(* IEC 61131-3 sources: plc-st-coding-agent/progress/evidence/f14_v10_full_20261113/jobs/codex_minimax-m27 (part 8) *)

(* ---- self-medium-03.raw_candidate_04.st ---- *)
TYPE EState :
    (
        IDLE    := 0,
        OPENING := 1,
        CLOSING := 2,
        FAULT   := 3
    )
END_TYPE

FUNCTION_BLOCK FB
VAR_INPUT
    openBtn    : BOOL;
    closeBtn   : BOOL;
    openLimit  : BOOL;
    closeLimit : BOOL;
    obstacle   : BOOL;
END_VAR
VAR_OUTPUT
    motorUp    : BOOL;
    motorDown  : BOOL;
    errorFlag  : BOOL;
END_VAR
VAR
    state          : EState := IDLE;
    prev_openBtn   : BOOL := FALSE;
    prev_closeBtn  : BOOL := FALSE;
    prev_obstacle  : BOOL := FALSE;
    openRTrig      : R_TRIG;
    closeRTrig     : R_TRIG;
    dualRTrig      : R_TRIG;
END_VAR

(*
ENGINEERING_CONTRACT
===================
| Output/State | Activation           | Retention           | Reset/Deactivation              | Scan Priority | Units   |
|--------------|----------------------|---------------------|----------------------------------|---------------|---------|
| motorUp      | IDLE+rising(openBtn) | Running continues   | obstacle/openLimit/FAULT         | Same-scan     | BOOL    |
| motorDown    | IDLE+rising(closeBtn)| Running continues   | obstacle/closeLimit/FAULT        | Same-scan     | BOOL    |
| errorFlag    | Any state+obstacle   | Latched in FAULT    | No obstacle+dualBtn rising edge  | Highest       | BOOL    |
| state=FAULT  | Any state+obstacle   | Until dualBtn reset | No obstacle+dualBtn rising edge  | Highest       | EState  |
| state=IDLE   | Power-on/limit/reset | Until rising edge   | -                                | Default       | EState  |
PUB001: power-on IDLE
PUB002: init FALSE
PUB003-005: no obstacle IDLE start (openBtn rising, closeBtn=FALSE, not openLimit)
PUB006: dual-btn does not start
PUB007: motor command same-scan on start
PUB008-009: button release / direction buttons ignored during movement
PUB010-011: limit stop same-scan, opposite limit irrelevant
PUB012: mutual exclusion always
PUB013-014: obstacle → both stop + FAULT (highest priority)
PUB017-018: errorFlag latched, motors stopped in FAULT
PUB019-021: reset requires no obstacle + dualBtn from not-both to both
PUB022-024: reset → IDLE, same-scan stop, then follow rule 1
*)

BEGIN
    openRTrig(CLK := openBtn);
    closeRTrig(CLK := closeBtn);
    dualRTrig(CLK := openBtn AND closeBtn);

    (* Priority 1: Obstacle → immediate both-stop + FAULT *)
    IF obstacle THEN
        motorUp   := FALSE;
        motorDown := FALSE;
        state     := FAULT;
        errorFlag := TRUE;
    ELSE
        CASE state OF
            IDLE:
                motorUp   := FALSE;
                motorDown := FALSE;
                (* Start opening: rising edge of openBtn, closeBtn=FALSE, not at openLimit *)
                IF openRTrig.Q AND NOT closeBtn AND NOT openLimit THEN
                    motorUp := TRUE;
                    state   := OPENING;
                (* Start closing: rising edge of closeBtn, openBtn=FALSE, not at closeLimit *)
                ELSIF closeRTrig.Q AND NOT openBtn AND NOT closeLimit THEN
                    motorDown := TRUE;
                    state     := CLOSING;
                END_IF;

            OPENING:
                motorUp   := TRUE;
                motorDown := FALSE;
                IF openLimit THEN
                    motorUp := FALSE;
                    state   := IDLE;
                END_IF;

            CLOSING:
                motorUp   := FALSE;
                motorDown := TRUE;
                IF closeLimit THEN
                    motorDown := FALSE;
                    state     := IDLE;
                END_IF;

            FAULT:
                motorUp   := FALSE;
                motorDown := FALSE;
                IF dualRTrig.Q THEN
                    errorFlag := FALSE;
                    state     := IDLE;
                END_IF;
        END_CASE;
    END_IF;

    prev_openBtn  := openBtn;
    prev_closeBtn := closeBtn;
    prev_obstacle := obstacle;
END_FUNCTION_BLOCK

(* CONTRACT_RULES [] *)

(* ---- self-medium-04.candidate_01.st ---- *)
(* ENGINEERING_CONTRACT
 * Filling Valve Controller - Discrete Scan State Machine
 *
 * | State            | Activation           | Retention           | Explicit Reset       | Same-scan Priority | Units/Boundaries     |
 * |------------------|----------------------|---------------------|----------------------|--------------------|----------------------|
 * | valveOpen=FALSE  | resetBtn rising      | N/A (output only)   | N/A                  | highest            | BOOL                 |
 * | valveOpen=TRUE   | rising(startBtn) & !prev(valveOpen) | while accVol < targetVol | resetBtn rising | 2nd            | accumulated REAL [0, ∞) |
 * | pendingFill=TRUE | valve closes (accVol>=target) | until doneSensor=TRUE OR new start OR reset | resetBtn rising | 3rd            | BOOL internal state       |
 * | fillsToday++     | doneSensor=TRUE & pendingFill | N/A (output only)  | resetBtn rising      | lowest             | INT [0..32767]           |
 *
 * PUB002: startBtn rising edge detection uses prevStartBtn
 * PUB003: resetBtn rising edge detection uses prevResetBtn
 * PUB004: doneSensor read as level each scan (PUB004)
 * PUB005: flowVol added each scan including start scan
 * PUB006: accumulated >= targetVol triggers valve close same scan
 * PUB007: doneSensor checked immediately after valve close
 * PUB008: if doneSensor=TRUE same scan, confirm and clear pendingFill
 * PUB009: if doneSensor=FALSE, pendingFill retained for later confirmation
 * PUB010: fillsToday increments by 1 per confirmation
 * PUB011: fillsToday saturates at 32767
 * PUB012: resetBtn rising clears all state (valveOpen, accumulatedVol, pendingFill, fillsToday)
 * PUB035: new start cancels pendingFill immediately
 * PUB043: continuous doneSensor=TRUE does not double-count
 *)
FUNCTION_BLOCK FB
VAR_INPUT
    startBtn    : BOOL;
    resetBtn    : BOOL;
    doneSensor  : BOOL;
    targetVol   : REAL;
    flowVol     : REAL;
END_VAR
VAR_OUTPUT
    valveOpen   : BOOL := FALSE;
    fillsToday  : INT  := 0;
END_VAR
VAR
    prevStartBtn    : BOOL := FALSE;
    prevResetBtn    : BOOL := FALSE;
    accumulatedVol  : REAL := 0.0;
    pendingFill     : BOOL := FALSE;
END_VAR

    // Priority 1: Reset clears everything, no other action this scan
    IF resetBtn AND NOT prevResetBtn THEN
        valveOpen       := FALSE;
        accumulatedVol  := 0.0;
        pendingFill     := FALSE;
        fillsToday      := 0;
        prevStartBtn    := startBtn;
        prevResetBtn    := resetBtn;
        RETURN;
    END_IF;

    // Priority 2: Start new bottle (clears any pending confirmation)
    IF startBtn AND NOT prevStartBtn THEN
        pendingFill    := FALSE;
        accumulatedVol := 0.0;
        valveOpen      := TRUE;
        // flowVol added in filling section below
    END_IF;

    // Priority 3: Filling state - accumulate flow and check target
    IF valveOpen THEN
        accumulatedVol := accumulatedVol + flowVol;
        IF accumulatedVol >= targetVol THEN
            valveOpen := FALSE;
            // Immediate doneSensor check after valve close
            IF doneSensor THEN
                pendingFill := FALSE;
                IF fillsToday < 32767 THEN
                    fillsToday := fillsToday + 1;
                END_IF;
            ELSE
                pendingFill := TRUE;
            END_IF;
        END_IF;
    END_IF;

    // Priority 4: Pending confirmation - wait for doneSensor
    IF pendingFill AND doneSensor THEN
        pendingFill := FALSE;
        IF fillsToday < 32767 THEN
            fillsToday := fillsToday + 1;
        END_IF;
    END_IF;

    prevStartBtn := startBtn;
    prevResetBtn := resetBtn;
END_FUNCTION_BLOCK

(* CONTRACT_RULES [] *)

(* ---- self-medium-04.raw_candidate_01.st ---- *)
(* ENGINEERING_CONTRACT
 * Filling Valve Controller - Discrete Scan State Machine
 *
 * | State            | Activation           | Retention           | Explicit Reset       | Same-scan Priority | Units/Boundaries     |
 * |------------------|----------------------|---------------------|----------------------|--------------------|----------------------|
 * | valveOpen=FALSE  | resetBtn rising      | N/A (output only)   | N/A                  | highest            | BOOL                 |
 * | valveOpen=TRUE   | rising(startBtn) & !prev(valveOpen) | while accVol < targetVol | resetBtn rising | 2nd            | accumulated REAL [0, ∞) |
 * | pendingFill=TRUE | valve closes (accVol>=target) | until doneSensor=TRUE OR new start OR reset | resetBtn rising | 3rd            | BOOL internal state       |
 * | fillsToday++     | doneSensor=TRUE & pendingFill | N/A (output only)  | resetBtn rising      | lowest             | INT [0..32767]           |
 *
 * PUB002: startBtn rising edge detection uses prevStartBtn
 * PUB003: resetBtn rising edge detection uses prevResetBtn
 * PUB004: doneSensor read as level each scan (PUB004)
 * PUB005: flowVol added each scan including start scan
 * PUB006: accumulated >= targetVol triggers valve close same scan
 * PUB007: doneSensor checked immediately after valve close
 * PUB008: if doneSensor=TRUE same scan, confirm and clear pendingFill
 * PUB009: if doneSensor=FALSE, pendingFill retained for later confirmation
 * PUB010: fillsToday increments by 1 per confirmation
 * PUB011: fillsToday saturates at 32767
 * PUB012: resetBtn rising clears all state (valveOpen, accumulatedVol, pendingFill, fillsToday)
 * PUB035: new start cancels pendingFill immediately
 * PUB043: continuous doneSensor=TRUE does not double-count
 *)
FUNCTION_BLOCK FB
VAR_INPUT
    startBtn    : BOOL;
    resetBtn    : BOOL;
    doneSensor  : BOOL;
    targetVol   : REAL;
    flowVol     : REAL;
END_VAR
VAR_OUTPUT
    valveOpen   : BOOL := FALSE;
    fillsToday  : INT  := 0;
END_VAR
VAR
    prevStartBtn    : BOOL := FALSE;
    prevResetBtn    : BOOL := FALSE;
    accumulatedVol  : REAL := 0.0;
    pendingFill     : BOOL := FALSE;
END_VAR

    // Priority 1: Reset clears everything, no other action this scan
    IF resetBtn AND NOT prevResetBtn THEN
        valveOpen       := FALSE;
        accumulatedVol  := 0.0;
        pendingFill     := FALSE;
        fillsToday      := 0;
        prevStartBtn    := startBtn;
        prevResetBtn    := resetBtn;
        RETURN;
    END_IF

    // Priority 2: Start new bottle (clears any pending confirmation)
    IF startBtn AND NOT prevStartBtn THEN
        pendingFill    := FALSE;
        accumulatedVol := 0.0;
        valveOpen      := TRUE;
        // flowVol added in filling section below
    END_IF

    // Priority 3: Filling state - accumulate flow and check target
    IF valveOpen THEN
        accumulatedVol := accumulatedVol + flowVol;
        IF accumulatedVol >= targetVol THEN
            valveOpen := FALSE;
            // Immediate doneSensor check after valve close
            IF doneSensor THEN
                pendingFill := FALSE;
                IF fillsToday < 32767 THEN
                    fillsToday := fillsToday + 1;
                END_IF
            ELSE
                pendingFill := TRUE;
            END_IF;
        END_IF;
    END_IF;

    // Priority 4: Pending confirmation - wait for doneSensor
    IF pendingFill AND doneSensor THEN
        pendingFill := FALSE;
        IF fillsToday < 32767 THEN
            fillsToday := fillsToday + 1;
        END_IF;
    END_IF;

    prevStartBtn := startBtn;
    prevResetBtn := resetBtn;
END_FUNCTION_BLOCK

(* CONTRACT_RULES [] *)

(* ---- self-medium-05.candidate_01.st ---- *)
FUNCTION_BLOCK FB
VAR_INPUT
    enable         : BOOL;
    resetBtn       : BOOL;
    scanSeconds    : LREAL;
    steamFlow      : LREAL;
    fuelFlow       : LREAL;
    steamTemp      : LREAL;
    steamPressure  : LREAL;
END_VAR
VAR_OUTPUT
    qualified      : BOOL;
    dataFault      : BOOL;
    qualifiedTon   : LREAL;
    fuelTon        : LREAL;
    revenue        : LREAL;
    cost           : LREAL;
    netProfit      : LREAL;
END_VAR
VAR
    prevResetBtn   : BOOL := FALSE;
    tmpFuelTon     : LREAL := 0.0;
    tmpQualifiedTon: LREAL := 0.0;
END_VAR

(* ENGINEERING_CONTRACT
 * PUB001-002:   enable=OFF → no accumulation; OFF+FAULT → freeze; reset rising → zero both immediately.
 * PUB003-004:   qualified = (steamTemp∈[447,453] ∧ steamPressure∈[3750,3850]) closed interval.
 * PUB005:       scanSeconds fault: ≤0.0 or >10.0 (10.0 itself is valid).
 * PUB006:       steamFlow fault: <0 or >90; fuelFlow fault: <0 or >6; negative values are faults.
 * PUB007-008:   Accumulation: fuelTon+=fuelFlow×scanSec/1000 when (enable ∧ ¬fault ∧ ¬resetRising).
 * PUB009-010:   Accumulation: qualifiedTon+=steamFlow×scanSec/1000 when (enable ∧ ¬fault ∧ qualified ∧ ¬resetRising).
 * PUB011:       Reset is edge-triggered; hold duration is irrelevant; one rising edge clears once.
 * PUB012-014:   Reset rising has highest priority; same-scan fault is reported but accumulators become 0.
 * PUB015-017:   revenue=qualifiedTon×280, cost=fuelTon×1500, netProfit=revenue−cost; updated every scan.
 * PUB018-022:   qualifiedTon, fuelTon, revenue, cost ≥0 always; netProfit may be negative.
 * Units:        steamFlow/fuelFlow in kg/s, scanSeconds in s → /1000 converts kg→t.
 *)

(* CONTRACT_RULES [] *)

qualified := (steamTemp >= 447.0) AND (steamTemp <= 453.0)
             AND (steamPressure >= 3750.0) AND (steamPressure <= 3850.0);

dataFault := (scanSeconds <= 0.0) OR (scanSeconds > 10.0)
             OR (steamFlow < 0.0) OR (steamFlow > 90.0)
             OR (fuelFlow < 0.0) OR (fuelFlow > 6.0);

IF resetBtn AND NOT prevResetBtn THEN
    tmpQualifiedTon := 0.0;
    tmpFuelTon := 0.0;
ELSE
    tmpQualifiedTon := qualifiedTon;
    tmpFuelTon := fuelTon;
    IF enable AND NOT dataFault THEN
        tmpFuelTon := fuelTon + fuelFlow * scanSeconds / 1000.0;
        IF qualified THEN
            tmpQualifiedTon := qualifiedTon + steamFlow * scanSeconds / 1000.0;
        END_IF;
    END_IF;
END_IF;

qualifiedTon := tmpQualifiedTon;
fuelTon      := tmpFuelTon;

revenue   := qualifiedTon * 280.0;
cost      := fuelTon * 1500.0;
netProfit := revenue - cost;

prevResetBtn := resetBtn;
END_FUNCTION_BLOCK

(* ---- self-medium-05.raw_candidate_01.st ---- *)
FUNCTION_BLOCK FB
VAR_INPUT
    enable         : BOOL;
    resetBtn       : BOOL;
    scanSeconds    : LREAL;
    steamFlow      : LREAL;
    fuelFlow       : LREAL;
    steamTemp      : LREAL;
    steamPressure  : LREAL;
END_VAR
VAR_OUTPUT
    qualified      : BOOL;
    dataFault      : BOOL;
    qualifiedTon   : LREAL;
    fuelTon        : LREAL;
    revenue        : LREAL;
    cost           : LREAL;
    netProfit      : LREAL;
END_VAR
VAR
    prevResetBtn   : BOOL := FALSE;
    tmpFuelTon     : LREAL := 0.0;
    tmpQualifiedTon: LREAL := 0.0;
END_VAR

(* ENGINEERING_CONTRACT
 * PUB001-002:   enable=OFF → no accumulation; OFF+FAULT → freeze; reset rising → zero both immediately.
 * PUB003-004:   qualified = (steamTemp∈[447,453] ∧ steamPressure∈[3750,3850]) closed interval.
 * PUB005:       scanSeconds fault: ≤0.0 or >10.0 (10.0 itself is valid).
 * PUB006:       steamFlow fault: <0 or >90; fuelFlow fault: <0 or >6; negative values are faults.
 * PUB007-008:   Accumulation: fuelTon+=fuelFlow×scanSec/1000 when (enable ∧ ¬fault ∧ ¬resetRising).
 * PUB009-010:   Accumulation: qualifiedTon+=steamFlow×scanSec/1000 when (enable ∧ ¬fault ∧ qualified ∧ ¬resetRising).
 * PUB011:       Reset is edge-triggered; hold duration is irrelevant; one rising edge clears once.
 * PUB012-014:   Reset rising has highest priority; same-scan fault is reported but accumulators become 0.
 * PUB015-017:   revenue=qualifiedTon×280, cost=fuelTon×1500, netProfit=revenue−cost; updated every scan.
 * PUB018-022:   qualifiedTon, fuelTon, revenue, cost ≥0 always; netProfit may be negative.
 * Units:        steamFlow/fuelFlow in kg/s, scanSeconds in s → /1000 converts kg→t.
 *)

(* CONTRACT_RULES [] *)

qualified := (steamTemp >= 447.0) AND (steamTemp <= 453.0)
             AND (steamPressure >= 3750.0) AND (steamPressure <= 3850.0);

dataFault := (scanSeconds <= 0.0) OR (scanSeconds > 10.0)
             OR (steamFlow < 0.0) OR (steamFlow > 90.0)
             OR (fuelFlow < 0.0) OR (fuelFlow > 6.0);

IF resetBtn AND NOT prevResetBtn THEN
    tmpQualifiedTon := 0.0;
    tmpFuelTon := 0.0;
ELSE
    tmpQualifiedTon := qualifiedTon;
    tmpFuelTon := fuelTon;
    IF enable AND NOT dataFault THEN
        tmpFuelTon := fuelTon + fuelFlow * scanSeconds / 1000.0;
        IF qualified THEN
            tmpQualifiedTon := qualifiedTon + steamFlow * scanSeconds / 1000.0;
        END_IF;
    END_IF;
END_IF;

qualifiedTon := tmpQualifiedTon;
fuelTon      := tmpFuelTon;

revenue   := qualifiedTon * 280.0;
cost      := fuelTon * 1500.0;
netProfit := revenue - cost;

prevResetBtn := resetBtn;
END_FUNCTION_BLOCK

(* ---- self-medium-06.candidate_01.st ---- *)
FUNCTION_BLOCK FB
VAR_INPUT
    enable         : BOOL;
    resetBtn       : BOOL;
    sensorValid    : BOOL;
    setpoint       : REAL;
    temperature    : REAL;
    scanSeconds    : REAL;
    bias           : REAL;
END_VAR
VAR_OUTPUT
    power          : REAL;
    correction     : REAL;
    fault          : BOOL;
END_VAR
VAR
    prevResetBtn   : BOOL := FALSE;
    prevEnable     : BOOL := FALSE;
    prevFault      : BOOL := FALSE;
    ePrev          : REAL := 0.0;
    historyCleared : BOOL := TRUE;
END_VAR

(* CONTRACT_RULES [] *)

(*
ENGINEERING_CONTRACT:
| Output/State  | Activation          | Retention       | Reset/Deactivation    | Same-Scan Priority | Units/Boundaries |
|---------------|---------------------|-----------------|-----------------------|--------------------|------------------|
| power         | enable & !fault     | Last valid      | !enable / fault /     | power=0 overrides  | 0..100 %         |
|               | & !resetRisingEdge  | clamp(bias+corr)| resetRisingEdge       | normal calc        |                  |
| correction    | enable & !fault     | Last valid      | !enable / fault /     | correction=0       | -30..30 %        |
|               | & !resetRisingEdge  | (no clamp)      | resetRisingEdge       | overrides calc     |                  |
| fault         | !sensorValid OR     | Latched while   | sensorValid & valid   | N/A (combinational)| BOOLEAN          |
|               | scanSeconds<=0/>10  | condition holds | scanSeconds           |                    |                  |
| ePrev         | Cleared on          | Holds across    | Cleared on !enable /  | N/A                | ℃               |
|               | first valid scan    | scans           | fault / resetRising   |                    |                  |
| historyCleared| Set TRUE on clear   | FALSE otherwise | Set TRUE on clear     | N/A                | BOOLEAN          |
| PUB001: enable controls autonomous mode
| PUB004: resetBtn is rising-edge command
| PUB006: fault triggers output zero + history clear
| PUB010: correction is centroid defuzzified
| PUB014: power = clamp(bias+correction, 0, 100)
*)
VAR
    resetRisingEdge : BOOL;
    e               : REAL;
    de              : REAL;
    x               : REAL;
    y               : REAL;
    muN_x           : REAL;
    muZ_x           : REAL;
    muP_x           : REAL;
    muN_y           : REAL;
    muZ_y           : REAL;
    muP_y           : REAL;
    wNN, wNZ, wNP   : REAL;
    wZN, wZZ, wZP   : REAL;
    wPN, wPZ, wPP   : REAL;
    sumW            : REAL;
    sumWc           : REAL;
END_VAR

// Fault detection (PUB006/PUB032)
fault := NOT sensorValid OR scanSeconds <= 0.0 OR scanSeconds > 10.0;

// Rising edge detection for resetBtn
resetRisingEdge := resetBtn AND NOT prevResetBtn;

// Clearing logic: first valid scan after disable/fault/reset rising edge
IF (!prevEnable OR resetRisingEdge OR prevFault) THEN
    power := 0.0;
    correction := 0.0;
    ePrev := 0.0;
    historyCleared := TRUE;
END_IF

// Main computation when enabled and not faulted
IF enable AND NOT fault THEN
    // Compute error (PUB001)
    e := setpoint - temperature;

    // Compute derivative (PUB002/PUB003)
    IF historyCleared THEN
        de := 0.0;
    ELSE
        de := (e - ePrev) / scanSeconds;
    END_IF

    // Normalize inputs (PUB005)
    x := LIMIT(-1.0, e / 10.0, 1.0);
    y := LIMIT(-1.0, de / 2.0, 1.0);

    // Membership functions (PUB004)
    muN_x := MAX(-x, 0.0);
    muZ_x := MAX(1.0 - ABS(x), 0.0);
    muP_x := MAX(x, 0.0);

    muN_y := MAX(-y, 0.0);
    muZ_y := MAX(1.0 - ABS(y), 0.0);
    muP_y := MAX(y, 0.0);

    // Rule weights: w(i,j) = mu_i(x) * mu_j(y)
    wNN := muN_x * muN_y;
    wNZ := muN_x * muZ_y;
    wNP := muN_x * muP_y;
    wZN := muZ_x * muN_y;
    wZZ := muZ_x * muZ_y;
    wZP := muZ_x * muP_y;
    wPN := muP_x * muN_y;
    wPZ := muP_x * muZ_y;
    wPP := muP_x * muP_y;

    // Centroid defuzzification (PUB010)
    sumW  := wNN + wNZ + wNP + wZN + wZZ + wZP + wPN + wPZ + wPP;
    sumWc := wNN * (-30.0) + wNZ * (-20.0) + wNP * (-10.0)
           + wZN * (-10.0) + wZZ * 0.0    + wZP * 10.0
           + wPN * 10.0   + wPZ * 20.0    + wPP * 30.0;

    IF sumW > 0.0 THEN
        correction := sumWc / sumW;
    ELSE
        correction := 0.0;
    END_IF

    // Output with clamping (PUB014)
    power := LIMIT(0.0, bias + correction, 100.0);

    // Update history for next scan
    ePrev := e;
    historyCleared := FALSE;
END_IF

// Update previous values for next scan
prevResetBtn := resetBtn;
prevEnable := enable;
prevFault := fault;
END_FUNCTION_BLOCK

(* ---- self-medium-06.candidate_02.st ---- *)
FUNCTION_BLOCK FB
VAR_INPUT
    enable         : BOOL;
    resetBtn       : BOOL;
    sensorValid    : BOOL;
    setpoint       : REAL;
    temperature    : REAL;
    scanSeconds    : REAL;
    bias           : REAL;
END_VAR
VAR_OUTPUT
    power          : REAL;
    correction     : REAL;
    fault          : BOOL;
END_VAR
VAR
    prevResetBtn   : BOOL := FALSE;
    prevEnable     : BOOL := FALSE;
    prevFault      : BOOL := FALSE;
    ePrev          : REAL := 0.0;
    historyCleared : BOOL := TRUE;
END_VAR

(* CONTRACT_RULES [] *)

(*
ENGINEERING_CONTRACT:
| Output/State  | Activation          | Retention       | Reset/Deactivation    | Same-Scan Priority | Units/Boundaries |
|---------------|---------------------|-----------------|-----------------------|--------------------|------------------|
| power         | enable & !fault     | Last valid      | !enable / fault /     | power=0 overrides  | 0..100 %         |
|               | & !resetRisingEdge  | clamp(bias+corr)| resetRisingEdge       | normal calc        |                  |
| correction    | enable & !fault     | Last valid      | !enable / fault /     | correction=0       | -30..30 %        |
|               | & !resetRisingEdge  | (no clamp)      | resetRisingEdge       | overrides calc     |                  |
| fault         | !sensorValid OR     | Latched while   | sensorValid & valid   | N/A (combinational)| BOOLEAN          |
|               | scanSeconds<=0/>10  | condition holds | scanSeconds           |                    |                  |
| ePrev         | Cleared on          | Holds across    | Cleared on !enable /  | N/A                | ℃               |
|               | first valid scan    | scans           | fault / resetRising   |                    |                  |
| historyCleared| Set TRUE on clear   | FALSE otherwise | Set TRUE on clear     | N/A                | BOOLEAN          |
| PUB001: enable controls autonomous mode
| PUB004: resetBtn is rising-edge command
| PUB006: fault triggers output zero + history clear
| PUB010: correction is centroid defuzzified
| PUB014: power = clamp(bias+correction, 0, 100)
*)
VAR
    resetRisingEdge : BOOL;
    e               : REAL;
    de              : REAL;
    x               : REAL;
    y               : REAL;
    muN_x           : REAL;
    muZ_x           : REAL;
    muP_x           : REAL;
    muN_y           : REAL;
    muZ_y           : REAL;
    muP_y           : REAL;
    wNN, wNZ, wNP   : REAL;
    wZN, wZZ, wZP   : REAL;
    wPN, wPZ, wPP   : REAL;
    sumW            : REAL;
    sumWc           : REAL;
END_VAR

// Fault detection (PUB006/PUB032)
fault := NOT sensorValid OR scanSeconds <= 0.0 OR scanSeconds > 10.0;

// Rising edge detection for resetBtn
resetRisingEdge := resetBtn AND NOT prevResetBtn;

// Clearing logic: first valid scan after disable/fault/reset rising edge
IF (NOT prevEnable OR resetRisingEdge OR prevFault) THEN
    power := 0.0;
    correction := 0.0;
    ePrev := 0.0;
    historyCleared := TRUE;
END_IF;

// Main computation when enabled and not faulted
IF enable AND NOT fault THEN
    // Compute error (PUB001)
    e := setpoint - temperature;

    // Compute derivative (PUB002/PUB003)
    IF historyCleared THEN
        de := 0.0;
    ELSE
        de := (e - ePrev) / scanSeconds;
    END_IF;

    // Normalize inputs (PUB005)
    x := LIMIT(-1.0, e / 10.0, 1.0);
    y := LIMIT(-1.0, de / 2.0, 1.0);

    // Membership functions (PUB004)
    muN_x := MAX(-x, 0.0);
    muZ_x := MAX(1.0 - ABS(x), 0.0);
    muP_x := MAX(x, 0.0);

    muN_y := MAX(-y, 0.0);
    muZ_y := MAX(1.0 - ABS(y), 0.0);
    muP_y := MAX(y, 0.0);

    // Rule weights: w(i,j) = mu_i(x) * mu_j(y)
    wNN := muN_x * muN_y;
    wNZ := muN_x * muZ_y;
    wNP := muN_x * muP_y;
    wZN := muZ_x * muN_y;
    wZZ := muZ_x * muZ_y;
    wZP := muZ_x * muP_y;
    wPN := muP_x * muN_y;
    wPZ := muP_x * muZ_y;
    wPP := muP_x * muP_y;

    // Centroid defuzzification (PUB010)
    sumW  := wNN + wNZ + wNP + wZN + wZZ + wZP + wPN + wPZ + wPP;
    sumWc := wNN * (-30.0) + wNZ * (-20.0) + wNP * (-10.0)
           + wZN * (-10.0) + wZZ * 0.0    + wZP * 10.0
           + wPN * 10.0   + wPZ * 20.0    + wPP * 30.0;

    IF sumW > 0.0 THEN
        correction := sumWc / sumW;
    ELSE
        correction := 0.0;
    END_IF;

    // Output with clamping (PUB014)
    power := LIMIT(0.0, bias + correction, 100.0);

    // Update history for next scan
    ePrev := e;
    historyCleared := FALSE;
END_IF;

// Update previous values for next scan
prevResetBtn := resetBtn;
prevEnable := enable;
prevFault := fault;
END_FUNCTION_BLOCK

(* ---- self-medium-06.raw_candidate_01.st ---- *)
FUNCTION_BLOCK FB
VAR_INPUT
    enable         : BOOL;
    resetBtn       : BOOL;
    sensorValid    : BOOL;
    setpoint       : REAL;
    temperature    : REAL;
    scanSeconds    : REAL;
    bias           : REAL;
END_VAR
VAR_OUTPUT
    power          : REAL;
    correction     : REAL;
    fault          : BOOL;
END_VAR
VAR
    prevResetBtn   : BOOL := FALSE;
    prevEnable     : BOOL := FALSE;
    prevFault      : BOOL := FALSE;
    ePrev          : REAL := 0.0;
    historyCleared : BOOL := TRUE;
END_VAR

(* CONTRACT_RULES [] *)

(*
ENGINEERING_CONTRACT:
| Output/State  | Activation          | Retention       | Reset/Deactivation    | Same-Scan Priority | Units/Boundaries |
|---------------|---------------------|-----------------|-----------------------|--------------------|------------------|
| power         | enable & !fault     | Last valid      | !enable / fault /     | power=0 overrides  | 0..100 %         |
|               | & !resetRisingEdge  | clamp(bias+corr)| resetRisingEdge       | normal calc        |                  |
| correction    | enable & !fault     | Last valid      | !enable / fault /     | correction=0       | -30..30 %        |
|               | & !resetRisingEdge  | (no clamp)      | resetRisingEdge       | overrides calc     |                  |
| fault         | !sensorValid OR     | Latched while   | sensorValid & valid   | N/A (combinational)| BOOLEAN          |
|               | scanSeconds<=0/>10  | condition holds | scanSeconds           |                    |                  |
| ePrev         | Cleared on          | Holds across    | Cleared on !enable /  | N/A                | ℃               |
|               | first valid scan    | scans           | fault / resetRising   |                    |                  |
| historyCleared| Set TRUE on clear   | FALSE otherwise | Set TRUE on clear     | N/A                | BOOLEAN          |
| PUB001: enable controls autonomous mode
| PUB004: resetBtn is rising-edge command
| PUB006: fault triggers output zero + history clear
| PUB010: correction is centroid defuzzified
| PUB014: power = clamp(bias+correction, 0, 100)
*)
VAR
    resetRisingEdge : BOOL;
    e               : REAL;
    de              : REAL;
    x               : REAL;
    y               : REAL;
    muN_x           : REAL;
    muZ_x           : REAL;
    muP_x           : REAL;
    muN_y           : REAL;
    muZ_y           : REAL;
    muP_y           : REAL;
    wNN, wNZ, wNP   : REAL;
    wZN, wZZ, wZP   : REAL;
    wPN, wPZ, wPP   : REAL;
    sumW            : REAL;
    sumWc           : REAL;
END_VAR

// Fault detection (PUB006/PUB032)
fault := NOT sensorValid OR scanSeconds <= 0.0 OR scanSeconds > 10.0;

// Rising edge detection for resetBtn
resetRisingEdge := resetBtn AND NOT prevResetBtn;

// Clearing logic: first valid scan after disable/fault/reset rising edge
IF (!prevEnable OR resetRisingEdge OR prevFault) THEN
    power := 0.0;
    correction := 0.0;
    ePrev := 0.0;
    historyCleared := TRUE;
END_IF

// Main computation when enabled and not faulted
IF enable AND NOT fault THEN
    // Compute error (PUB001)
    e := setpoint - temperature;

    // Compute derivative (PUB002/PUB003)
    IF historyCleared THEN
        de := 0.0;
    ELSE
        de := (e - ePrev) / scanSeconds;
    END_IF

    // Normalize inputs (PUB005)
    x := LIMIT(-1.0, e / 10.0, 1.0);
    y := LIMIT(-1.0, de / 2.0, 1.0);

    // Membership functions (PUB004)
    muN_x := MAX(-x, 0.0);
    muZ_x := MAX(1.0 - ABS(x), 0.0);
    muP_x := MAX(x, 0.0);

    muN_y := MAX(-y, 0.0);
    muZ_y := MAX(1.0 - ABS(y), 0.0);
    muP_y := MAX(y, 0.0);

    // Rule weights: w(i,j) = mu_i(x) * mu_j(y)
    wNN := muN_x * muN_y;
    wNZ := muN_x * muZ_y;
    wNP := muN_x * muP_y;
    wZN := muZ_x * muN_y;
    wZZ := muZ_x * muZ_y;
    wZP := muZ_x * muP_y;
    wPN := muP_x * muN_y;
    wPZ := muP_x * muZ_y;
    wPP := muP_x * muP_y;

    // Centroid defuzzification (PUB010)
    sumW  := wNN + wNZ + wNP + wZN + wZZ + wZP + wPN + wPZ + wPP;
    sumWc := wNN * (-30.0) + wNZ * (-20.0) + wNP * (-10.0)
           + wZN * (-10.0) + wZZ * 0.0    + wZP * 10.0
           + wPN * 10.0   + wPZ * 20.0    + wPP * 30.0;

    IF sumW > 0.0 THEN
        correction := sumWc / sumW;
    ELSE
        correction := 0.0;
    END_IF

    // Output with clamping (PUB014)
    power := LIMIT(0.0, bias + correction, 100.0);

    // Update history for next scan
    ePrev := e;
    historyCleared := FALSE;
END_IF

// Update previous values for next scan
prevResetBtn := resetBtn;
prevEnable := enable;
prevFault := fault;
END_FUNCTION_BLOCK

(* ---- self-medium-06.raw_candidate_02.st ---- *)
FUNCTION_BLOCK FB
VAR_INPUT
    enable         : BOOL;
    resetBtn       : BOOL;
    sensorValid    : BOOL;
    setpoint       : REAL;
    temperature    : REAL;
    scanSeconds    : REAL;
    bias           : REAL;
END_VAR
VAR_OUTPUT
    power          : REAL;
    correction     : REAL;
    fault          : BOOL;
END_VAR
VAR
    prevResetBtn   : BOOL := FALSE;
    prevEnable     : BOOL := FALSE;
    prevFault      : BOOL := FALSE;
    ePrev          : REAL := 0.0;
    historyCleared : BOOL := TRUE;
END_VAR

(* CONTRACT_RULES [] *)

(*
ENGINEERING_CONTRACT:
| Output/State  | Activation          | Retention       | Reset/Deactivation    | Same-Scan Priority | Units/Boundaries |
|---------------|---------------------|-----------------|-----------------------|--------------------|------------------|
| power         | enable & !fault     | Last valid      | !enable / fault /     | power=0 overrides  | 0..100 %         |
|               | & !resetRisingEdge  | clamp(bias+corr)| resetRisingEdge       | normal calc        |                  |
| correction    | enable & !fault     | Last valid      | !enable / fault /     | correction=0       | -30..30 %        |
|               | & !resetRisingEdge  | (no clamp)      | resetRisingEdge       | overrides calc     |                  |
| fault         | !sensorValid OR     | Latched while   | sensorValid & valid   | N/A (combinational)| BOOLEAN          |
|               | scanSeconds<=0/>10  | condition holds | scanSeconds           |                    |                  |
| ePrev         | Cleared on          | Holds across    | Cleared on !enable /  | N/A                | ℃               |
|               | first valid scan    | scans           | fault / resetRising   |                    |                  |
| historyCleared| Set TRUE on clear   | FALSE otherwise | Set TRUE on clear     | N/A                | BOOLEAN          |
| PUB001: enable controls autonomous mode
| PUB004: resetBtn is rising-edge command
| PUB006: fault triggers output zero + history clear
| PUB010: correction is centroid defuzzified
| PUB014: power = clamp(bias+correction, 0, 100)
*)
VAR
    resetRisingEdge : BOOL;
    e               : REAL;
    de              : REAL;
    x               : REAL;
    y               : REAL;
    muN_x           : REAL;
    muZ_x           : REAL;
    muP_x           : REAL;
    muN_y           : REAL;
    muZ_y           : REAL;
    muP_y           : REAL;
    wNN, wNZ, wNP   : REAL;
    wZN, wZZ, wZP   : REAL;
    wPN, wPZ, wPP   : REAL;
    sumW            : REAL;
    sumWc           : REAL;
END_VAR

// Fault detection (PUB006/PUB032)
fault := NOT sensorValid OR scanSeconds <= 0.0 OR scanSeconds > 10.0;

// Rising edge detection for resetBtn
resetRisingEdge := resetBtn AND NOT prevResetBtn;

// Clearing logic: first valid scan after disable/fault/reset rising edge
IF (NOT prevEnable OR resetRisingEdge OR prevFault) THEN
    power := 0.0;
    correction := 0.0;
    ePrev := 0.0;
    historyCleared := TRUE;
END_IF

// Main computation when enabled and not faulted
IF enable AND NOT fault THEN
    // Compute error (PUB001)
    e := setpoint - temperature;

    // Compute derivative (PUB002/PUB003)
    IF historyCleared THEN
        de := 0.0;
    ELSE
        de := (e - ePrev) / scanSeconds;
    END_IF

    // Normalize inputs (PUB005)
    x := LIMIT(-1.0, e / 10.0, 1.0);
    y := LIMIT(-1.0, de / 2.0, 1.0);

    // Membership functions (PUB004)
    muN_x := MAX(-x, 0.0);
    muZ_x := MAX(1.0 - ABS(x), 0.0);
    muP_x := MAX(x, 0.0);

    muN_y := MAX(-y, 0.0);
    muZ_y := MAX(1.0 - ABS(y), 0.0);
    muP_y := MAX(y, 0.0);

    // Rule weights: w(i,j) = mu_i(x) * mu_j(y)
    wNN := muN_x * muN_y;
    wNZ := muN_x * muZ_y;
    wNP := muN_x * muP_y;
    wZN := muZ_x * muN_y;
    wZZ := muZ_x * muZ_y;
    wZP := muZ_x * muP_y;
    wPN := muP_x * muN_y;
    wPZ := muP_x * muZ_y;
    wPP := muP_x * muP_y;

    // Centroid defuzzification (PUB010)
    sumW  := wNN + wNZ + wNP + wZN + wZZ + wZP + wPN + wPZ + wPP;
    sumWc := wNN * (-30.0) + wNZ * (-20.0) + wNP * (-10.0)
           + wZN * (-10.0) + wZZ * 0.0    + wZP * 10.0
           + wPN * 10.0   + wPZ * 20.0    + wPP * 30.0;

    IF sumW > 0.0 THEN
        correction := sumWc / sumW;
    ELSE
        correction := 0.0;
    END_IF

    // Output with clamping (PUB014)
    power := LIMIT(0.0, bias + correction, 100.0);

    // Update history for next scan
    ePrev := e;
    historyCleared := FALSE;
END_IF

// Update previous values for next scan
prevResetBtn := resetBtn;
prevEnable := enable;
prevFault := fault;
END_FUNCTION_BLOCK

(* ---- public-medium-08.candidate_03.st ---- *)
Looking at the test case `"1..2.3"` producing `16777731` (0x01000203 = "1.0.2.3"), the issue is clear: the original implementation treats consecutive dots as a separator followed by an empty segment (defaulting to 0), which violates PUB003 ("nondigit segment" should produce 0).

The fix requires tracking whether the previous character was a separator so consecutive dots are rejected as malformed input.
[TOOL_CALL]
{tool => "apply_patch", args => {
  --path "E:\PLC_Dev\evidence\real_experiments\f14_v10_full_20261113\cli_private\ee35760ddffe45d99850d3a9dd357ba5\IPv4_Parse.st"
  --patch "*** Begin Patch\n*** Update File: E:\\PLC_Dev\\evidence\\real_experiments\\f14_v10_full_20261113\\cli_private\\ee35760ddffe45d99850d3a9dd357ba5\\IPv4_Parse.st\n@@ \n (* ENGINEERING_CONTRACT\n   PUB001: Parse dotted-decimal IPv4, validate 4 numeric segments 0-255\n   PUB002: Network byte order assembly (MSB=first segment)\n   PUB003: Invalid input → ipValue=0 (malformed, nondigit, wrong count, OOR)\n   PUB004: Valid 0.0.0.0 also produces 0 (by assembly)\n   \n   State retention: None (stateless function block)\n   Reset behavior: None (no reset input specified)\n   First scan: Same as subsequent (no edge memory)\n*)\n\n(* CONTRACT_RULES [] *)\n\nFUNCTION_BLOCK IPv4_Parse\nVAR_INPUT\n    ipText : STRING(254);\nEND_VAR\nVAR_OUTPUT\n    ipValue : UDINT := 0;\nEND_VAR\nVAR\n    tmp_pos : UDINT;\n    tmp_seg_idx : UDINT;\n    tmp_char : BYTE;\n    tmp_seg_val : UDINT;\n    tmp_result : UDINT;\n    tmp_prev_was_sep : BOOL;\n    tmp_digit_accumulated : BOOL;\nEND_VAR\n\ntmp_pos := 0;\ntmp_seg_idx := 0;\ntmp_result := 0;\ntmp_seg_val := 0;\ntmp_prev_was_sep := FALSE;\ntmp_digit_accumulated := FALSE;\n\nWHILE tmp_pos < LEN(ipText) DO\n    tmp_char := ipText[tmp_pos];\n    \n    IF tmp_char >= 48 AND tmp_char <= 57 THEN\n        tmp_seg_val := tmp_seg_val * 10 + TO_UDINT(tmp_char - 48);\n        \n        IF tmp_seg_val > 255 THEN\n            ipValue := 0;\n            RETURN;\n        END_IF;\n        \n        tmp_digit_accumulated := TRUE;\n        tmp_prev_was_sep := FALSE;\n        tmp_pos := tmp_pos + 1;\n        \n    ELSIF tmp_char = 46 THEN\n        // Separator: reject if leading, trailing, or consecutive\n        IF tmp_prev_was_sep OR NOT tmp_digit_accumulated THEN\n            ipValue := 0;\n            RETURN;\n        END_IF;\n        \n        IF tmp_seg_idx >= 3 THEN\n            ipValue := 0;\n            RETURN;\n        END_IF;\n        \n        CASE tmp_seg_idx OF\n            0: tmp_result := SHL(tmp_seg_val, 24);\n            1: tmp_result := tmp_result OR SHL(tmp_seg_val, 16);\n            2: tmp_result := tmp_result OR SHL(tmp_seg_val, 8);\n            3: tmp_result := tmp_result OR tmp_seg_val;\n        END_CASE;\n        \n        tmp_seg_idx := tmp_seg_idx + 1;\n        tmp_seg_val := 0;\n        tmp_prev_was_sep := TRUE;\n        tmp_digit_accumulated := FALSE;\n        tmp_pos := tmp_pos + 1;\n        \n    ELSE\n        ipValue := 0;\n        RETURN;\n    END_IF;\nEND_WHILE;\n\n// Reject trailing separator\nIF tmp_prev_was_sep OR NOT tmp_digit_accumulated THEN\n    ipValue := 0;\n    RETURN;\nEND_IF;\n\nIF tmp_seg_idx <> 3 THEN\n    ipValue := 0;\nELSE\n    tmp_result := tmp_result OR tmp_seg_val;\n    ipValue := tmp_result;\nEND_IF;\n\nEND_FUNCTION_BLOCK"
}}
[/TOOL_CALL]

(* ---- public-medium-08.raw_candidate_03.st ---- *)
Looking at the test case `"1..2.3"` producing `16777731` (0x01000203 = "1.0.2.3"), the issue is clear: the original implementation treats consecutive dots as a separator followed by an empty segment (defaulting to 0), which violates PUB003 ("nondigit segment" should produce 0).

The fix requires tracking whether the previous character was a separator so consecutive dots are rejected as malformed input.
[TOOL_CALL]
{tool => "apply_patch", args => {
  --path "E:\PLC_Dev\evidence\real_experiments\f14_v10_full_20261113\cli_private\ee35760ddffe45d99850d3a9dd357ba5\IPv4_Parse.st"
  --patch "*** Begin Patch\n*** Update File: E:\\PLC_Dev\\evidence\\real_experiments\\f14_v10_full_20261113\\cli_private\\ee35760ddffe45d99850d3a9dd357ba5\\IPv4_Parse.st\n@@ \n (* ENGINEERING_CONTRACT\n   PUB001: Parse dotted-decimal IPv4, validate 4 numeric segments 0-255\n   PUB002: Network byte order assembly (MSB=first segment)\n   PUB003: Invalid input → ipValue=0 (malformed, nondigit, wrong count, OOR)\n   PUB004: Valid 0.0.0.0 also produces 0 (by assembly)\n   \n   State retention: None (stateless function block)\n   Reset behavior: None (no reset input specified)\n   First scan: Same as subsequent (no edge memory)\n*)\n\n(* CONTRACT_RULES [] *)\n\nFUNCTION_BLOCK IPv4_Parse\nVAR_INPUT\n    ipText : STRING(254);\nEND_VAR\nVAR_OUTPUT\n    ipValue : UDINT := 0;\nEND_VAR\nVAR\n    tmp_pos : UDINT;\n    tmp_seg_idx : UDINT;\n    tmp_char : BYTE;\n    tmp_seg_val : UDINT;\n    tmp_result : UDINT;\n    tmp_prev_was_sep : BOOL;\n    tmp_digit_accumulated : BOOL;\nEND_VAR\n\ntmp_pos := 0;\ntmp_seg_idx := 0;\ntmp_result := 0;\ntmp_seg_val := 0;\ntmp_prev_was_sep := FALSE;\ntmp_digit_accumulated := FALSE;\n\nWHILE tmp_pos < LEN(ipText) DO\n    tmp_char := ipText[tmp_pos];\n    \n    IF tmp_char >= 48 AND tmp_char <= 57 THEN\n        tmp_seg_val := tmp_seg_val * 10 + TO_UDINT(tmp_char - 48);\n        \n        IF tmp_seg_val > 255 THEN\n            ipValue := 0;\n            RETURN;\n        END_IF;\n        \n        tmp_digit_accumulated := TRUE;\n        tmp_prev_was_sep := FALSE;\n        tmp_pos := tmp_pos + 1;\n        \n    ELSIF tmp_char = 46 THEN\n        // Separator: reject if leading, trailing, or consecutive\n        IF tmp_prev_was_sep OR NOT tmp_digit_accumulated THEN\n            ipValue := 0;\n            RETURN;\n        END_IF;\n        \n        IF tmp_seg_idx >= 3 THEN\n            ipValue := 0;\n            RETURN;\n        END_IF;\n        \n        CASE tmp_seg_idx OF\n            0: tmp_result := SHL(tmp_seg_val, 24);\n            1: tmp_result := tmp_result OR SHL(tmp_seg_val, 16);\n            2: tmp_result := tmp_result OR SHL(tmp_seg_val, 8);\n            3: tmp_result := tmp_result OR tmp_seg_val;\n        END_CASE;\n        \n        tmp_seg_idx := tmp_seg_idx + 1;\n        tmp_seg_val := 0;\n        tmp_prev_was_sep := TRUE;\n        tmp_digit_accumulated := FALSE;\n        tmp_pos := tmp_pos + 1;\n        \n    ELSE\n        ipValue := 0;\n        RETURN;\n    END_IF;\nEND_WHILE;\n\n// Reject trailing separator\nIF tmp_prev_was_sep OR NOT tmp_digit_accumulated THEN\n    ipValue := 0;\n    RETURN;\nEND_IF;\n\nIF tmp_seg_idx <> 3 THEN\n    ipValue := 0;\nELSE\n    tmp_result := tmp_result OR tmp_seg_val;\n    ipValue := tmp_result;\nEND_IF;\n\nEND_FUNCTION_BLOCK"
}}
[/TOOL_CALL]
